// TwinCAT 3 PLC project UnitTest
// ProgramVersion: 3.1.4026.29
// libraries:
//   [SampleLib], * (MyCompany)
//   Tc2_Standard, * (Beckhoff Automation GmbH)
//   Tc2_System, * (Beckhoff Automation GmbH)
//   Tc3_PlcTestFramework, * (Beckhoff Automation GmbH)
// project tree:
//   / PlcTask.TcTTO
//   POUs/ MAIN.TcPOU
//   TestCases/ FB_TestSum.TcPOU, FB_TestDiff.TcPOU, FB_TestProd.TcPOU, FB_TestDiv.TcPOU
// (motion and I/O tree: see PLC project mylib)
// real-time tasks:
//   TASK PlcTask: cycle T#10ms, priority 20, ADS port 350
//   TASK PlcTask1: cycle T#10ms, priority 21, ADS port 351

CONFIGURATION UnitTest
    RESOURCE PLC ON TwinCAT3
        TASK PlcTask(INTERVAL := T#10ms, PRIORITY := 21);
        PROGRAM MAIN WITH PlcTask : MAIN;
    END_RESOURCE
END_CONFIGURATION

// ---- POUs/MAIN.TcPOU
PROGRAM MAIN
VAR
	//instantiation of the test case function blocks
	fbT1	: FB_TestSum;   //Test case for the FB_Sum function block from the library
	fbT2	: FB_TestDiff;  //Test case for the FB_Diff function block from the library
	fbT3	: FB_TestProd;  //Test case for the FB_Prod function block from the library
	fbT4	: FB_TestDiv;   //Test case for the FB_Div function block from the library
END_VAR

//To have the source code for a library’s unit tests directly within the same solution, it is advisable to enable the option “Allow the project to be referenced as a library” in the library project. This option makes it possible to run the tests at any time without having to install the library on the system. It is therefore particularly useful for use in CI/CD pipelines, as the command to install the libraries does not need to be executed.

// Calling the TestController (which is located in the library and acts as the interface to the clients) 
Tc3_PlcTestFramework.F_CallTestController();

END_PROGRAM

// ---- TestCases/FB_TestSum.TcPOU
{ attribute 'Name':='TB_Sum-Test' }
{ attribute 'Timeout':='t#20s' }
{ attribute 'Owner':='TestOwner' }
{ attribute 'Category':='Math/addition and subtraction' }
FUNCTION_BLOCK FB_TestSum EXTENDS FB_TestCaseBase
VAR_INPUT
END_VAR
VAR_OUTPUT
END_VAR
VAR
	myFB : SampleLib.FB_Sum;    // instance of the function block to be tested
	expectedValue : UINT;       // value to be expected from this test
	result: UINT;				// calculated value, actual result of the function block call
END_VAR

// can of the function block to execute the test: in this casae 2 + 2 = 4
myFB(var1:= 2, var2:= 2, result=> result);

// Explicit assignment of the expected value, as the comparison is performed using the “any” data type
expectedValue:=4;

// Check the result against the expected value; if it does not match, the error message passed here is displayed
AssertEqual(anyActual:= result, anyExpected:= expectedValue, sMessage:= 'Addition with the FB_Sum function block is incorrect!');

// in the event that the result of the comparison matches, confirmation that the test case was successful and that no further tests will be carried out in this function block
Succeed();

//Must be implemented if you want to use fastmode
METHOD CleanUp : BOOL
CleanUp:=true;
END_METHOD

END_FUNCTION_BLOCK

// ---- TestCases/FB_TestDiff.TcPOU
{ attribute 'Name':='FB_Diff-Test' }
{ attribute 'Timeout':='t#20s' }
{ attribute 'Owner':='TestOwner' }
{ attribute 'Category':='Math/addition and subtraction' }
FUNCTION_BLOCK FB_TestDiff EXTENDS FB_TestCaseBase
VAR_INPUT
END_VAR
VAR_OUTPUT
END_VAR
VAR
	myFB : SampleLib.FB_Diff;   // instance of the function block to be tested
	expectedValue : UINT;       // value to be expected from this test
	result: UINT;				// calculated value, actual result of the function block call
END_VAR

// can of the function block to execute the test: 4 - 2 = 2
myFB(var1:= 4, var2:= 2, result=> result);

// Explicit assignment of the expected value, as the comparison is performed using the “any” data type
expectedValue:=2;

// Check the result against the expected value; if it does not match, the error message passed here is displayed
AssertEqual(anyActual:= result, anyExpected:= expectedValue, sMessage:= 'Subtraction with the FB_Diff function block is incorrect!');

// in the event that the result of the comparison matches, confirmation that the test case was successful and that no further tests will be carried out in this function block
Succeed();

//Must be implemented if you want to use fastmode
METHOD CleanUp : BOOL
CleanUp:=true;
END_METHOD

END_FUNCTION_BLOCK

// ---- TestCases/FB_TestProd.TcPOU
{ attribute 'Name':='TB_Prod-Test' }
{ attribute 'Timeout':='t#20s' }
{ attribute 'Owner':='TestOwner' }
{ attribute 'Category':='Math/multiplication and division ' }
FUNCTION_BLOCK FB_TestProd EXTENDS FB_TestCaseBase
VAR_INPUT
END_VAR
VAR_OUTPUT
END_VAR
VAR
	myFB : SampleLib.FB_Prod;   // instance of the function block to be tested
	expectedValue : UINT;       // value to be expected from this test
	result: UINT;				// calculated value, actual result of the function block call
END_VAR

// can of the function block to execute the test: 2 * 2 = 4
myFB(var1:= 2, var2:= 2, result=> result);

// Explicit assignment of the expected value, as the comparison is performed using the “any” data type
expectedValue:=4;

// Check the result against the expected value; if it does not match, the error message passed here is displayed
AssertEqual(anyActual:= result, anyExpected:= expectedValue, sMessage:= 'Multiplication with the FB_Prod function block is incorrect!');

// in the event that the result of the comparison matches, confirmation that the test case was successful and that no further tests will be carried out in this function block
Succeed();

//Must be implemented if you want to use fastmode
METHOD CleanUp : BOOL
CleanUp:=true;
END_METHOD

END_FUNCTION_BLOCK

// ---- TestCases/FB_TestDiv.TcPOU
{ attribute 'Name':='TB_Div-Test' }
{ attribute 'Timeout':='t#20s' }
{ attribute 'Owner':='TestOwner' }
{ attribute 'Category':='Math/multiplication and division ' }
FUNCTION_BLOCK FB_TestDiv EXTENDS FB_TestCaseBase
VAR_INPUT
END_VAR
VAR_OUTPUT
END_VAR
VAR
	myFB : SampleLib.FB_Div;    // instance of the function block to be tested
	expectedValue : UINT;       // value to be expected from this test
	result: UINT;				// calculated value, actual result of the function block call
END_VAR

// can of the function block to execute the test: 8 / 2 = 4
myFB(var1:= 8, var2:= 2, result=> result);

// Explicit assignment of the expected value, as the comparison is performed using the “any” data type
expectedValue:=4;

// Check the result against the expected value; if it does not match, the error message passed here is displayed
AssertEqual(anyActual:= result, anyExpected:= expectedValue, sMessage:= 'Division with the FB_Div function block is incorrect!');

// in the event that the result of the comparison matches, confirmation that the test case was successful and that no further tests will be carried out in this function block
Succeed();

//Must be implemented if you want to use fastmode
METHOD CleanUp : BOOL
CleanUp:=true;
END_METHOD

END_FUNCTION_BLOCK
